(* Arrival Time Monitor core, an abstract base by convention: thin ND-framework
   state-mover wrapper that holds only references, interfaces and the shared
   sub-FBs. The state bridge is here as REFERENCE TO UINT (eEnumSetRef and
   eEnumGetRef) and the body runs on it, but the enum variables, the state
   storage and the state names belong to the derived type, which passes them
   in. Y mover via FB_PositionStatePMPSND over one motor, plus a
   tick site for the in-beam thermocouple and flow meter.

   A derived type supplies everything that depends on the state list:
     - eEnumSet and eEnumGet, the device enum (UINT base, OUT = 1, then the
       targets) with the MMS:STATE:SET and MMS:STATE:GET pytmc pragmas, so the
       EPICS state menu comes from that enum;
     - afbStateDefaults, one FB_CC_InternalStateConfig per state, which writes
       the per-state sName and fDelta;
     - an FB_Init that repeats the inputs below and binds eEnumSetRef and
       eEnumGetRef to the enum variables, and a CallAfterInit that calls the
       configurators. The base CallAfterInit runs on its own through the
       call_after_init attribute.
   FB_ATM is the library derived type (E_ATM_States). A device with another
   state list derives this FB the same way.

   State 1 is OUT, which vetoes the thermocouple. *)
{attribute 'call_after_init'}
FUNCTION_BLOCK FB_ATM_Core
VAR
    {attribute 'pytmc' := 'pv: STC:01'}
    fbTempSensor1 : FB_CC_TempSensor;

    {attribute 'pytmc' := 'pv: FWM'}
    fbFlowMeter : FB_AnalogInput := (iTermBits := 15, fTermMax := 60, fTermMin := 0);

    {attribute 'no_copy'}
    aiMotionStage         : REFERENCE TO ARRAY[1..MotionConstants.MAX_STATE_MOTORS] OF I_MotionStage;
    {attribute 'no_copy'}
    astPositionState      : REFERENCE TO ARRAY[1..MotionConstants.MAX_STATE_MOTORS]
                                            OF ARRAY[1..GeneralConstants.MAX_STATES] OF ST_PositionState;
    {attribute 'no_copy'}
    fbFFHWO               : REFERENCE TO FB_HardwareFFOutput;
    {attribute 'no_copy'}
    fbArbiter             : REFERENCE TO FB_Arbiter;
    sDeviceName           : STRING;
    sTransitionKey        : STRING;
    bEnableMotion         : BOOL := TRUE;
    bEnableBeamParams     : BOOL;
    bEnablePositionLimits : BOOL;
    bReadDBNow            : BOOL;
    bFileReaderBusy       : REFERENCE TO BOOL;
    bFileReaderError      : REFERENCE TO BOOL;

    {attribute 'no_copy'}
    eEnumSetRef           : REFERENCE TO UINT;
    {attribute 'no_copy'}
    eEnumGetRef           : REFERENCE TO UINT;

    {attribute 'pytmc' := 'pv: MMS'}
    fbStates : FB_PositionStatePMPSND(
        aiMotionStage         := aiMotionStage,
        astPositionState      := astPositionState,
        nActiveMotorCount     := nStateMotorCount,
        eEnumSet              := eEnumSetRef,
        eEnumGet              := eEnumGetRef,
        bEnableMotion         := bEnableMotion,
        eMotionRequestPolicy  := E_MotionRequestPolicy.INTERRUPT,
        bEnableBeamParams     := bEnableBeamParams,
        bEnablePositionLimits := bEnablePositionLimits,
        bReadDBNow            := bReadDBNow,
        bFileReaderBusy       := bFileReaderBusy,
        bFileReaderError      := bFileReaderError,
        fbFFHWO               := fbFFHWO,
        fbArbiter             := fbArbiter,
        sDeviceName           := sDeviceName,
        sTransitionKey        := sTransitionKey
    );
END_VAR
VAR_OUTPUT
    // The PMPS database lookup associated with the current position state.
    stDbStateParams: ST_DbStateParams;
END_VAR
VAR CONSTANT
    (* Number of motors the state mover drives. Every device here has one state
       motor, in slot 1; the code around fbStates assumes it. *)
    nStateMotorCount : UINT := 1;
    (* ATM-wide default tolerance for state in-position detection. Derived
       types pass it to their afbStateDefaults. *)
    FDELTA_DEFAULT : LREAL := 2;
    // State value of OUT in every ATM enum.
    nOutState : UINT := 1;
END_VAR

IF NOT __ISVALIDREF(aiMotionStage)
   OR NOT __ISVALIDREF(astPositionState)
   OR NOT __ISVALIDREF(fbFFHWO)
   OR NOT __ISVALIDREF(fbArbiter)
   OR NOT __ISVALIDREF(eEnumSetRef)
   OR NOT __ISVALIDREF(eEnumGetRef) THEN
    RETURN;
END_IF

fbStates(
    stDbStateParams => stDbStateParams
);

// Faults only while something is in the beam (not OUT).
fbTempSensor1(
    fFaultThreshold := fbStates.stDbStateParams.stReactiveParams.nTempSP,
    bVeto           := eEnumGetRef = nOutState,
    sDevName        := sDeviceName,
    io_fbFFHWO      := fbFFHWO
);

fbFlowMeter();

(* Auto-fired after FB_Init. Wires fbStates through CallAfterInitCore. *)
{attribute 'call_after_init'}
METHOD CallAfterInit
THIS^.CallAfterInitCore();
END_METHOD

(* Wires fbStates with the references this FB holds, through
   CallAfterInitStateMover / CallAfterInitPMPS, because fbStates' inline-init
   ran first and forwarded nil refs. Does nothing while the essential refs are
   still nil. CallAfterInit calls it. A derived type that was re-wired after its
   host FB's CallAfterInit calls it again through SUPER^. *)
METHOD CallAfterInitCore
IF NOT __ISVALIDREF(aiMotionStage)
   OR NOT __ISVALIDREF(astPositionState)
   OR NOT __ISVALIDREF(eEnumSetRef)
   OR NOT __ISVALIDREF(eEnumGetRef) THEN
    RETURN;
END_IF

THIS^.fbStates.CallAfterInitStateMover(
    aiMotionStage         := aiMotionStage,
    astPositionState      := astPositionState,
    nActiveMotorCount     := nStateMotorCount,
    eEnumSet              := eEnumSetRef,
    eEnumGet              := eEnumGetRef,
    bEnableMotion         := bEnableMotion,
    eMotionRequestPolicy  := E_MotionRequestPolicy.INTERRUPT,
);

THIS^.fbStates.CallAfterInitPMPS(
    aiMotionStage         := aiMotionStage,
    astPositionState      := astPositionState,
    bEnableBeamParams     := bEnableBeamParams,
    bEnablePositionLimits := bEnablePositionLimits,
    bReadDBNow            := bReadDBNow,
    bFileReaderBusy       := bFileReaderBusy,
    bFileReaderError      := bFileReaderError,
    fbFFHWO               := fbFFHWO,
    fbArbiter             := fbArbiter,
    sDeviceName           := sDeviceName,
    sTransitionKey        := sTransitionKey
);
END_METHOD

(* Stores FB_Init inputs into instance fields; every non-value input is
   REFERENCE TO, REF= bound for the FB lifetime. fbStates inline-init
   captured these params at construction, so this records the same refs
   on THIS^ for body use and live caller writes. *)
{attribute 'analysis' := '-33'}
METHOD FB_Init : BOOL
VAR_INPUT
    bInitRetains           : BOOL;
    bInCopyCode            : BOOL;
    aiMotionStage          : REFERENCE TO ARRAY[1..MotionConstants.MAX_STATE_MOTORS] OF I_MotionStage;
    astPositionState       : REFERENCE TO ARRAY[1..MotionConstants.MAX_STATE_MOTORS]
                                            OF ARRAY[1..GeneralConstants.MAX_STATES] OF ST_PositionState;
    fbFFHWO                : REFERENCE TO FB_HardwareFFOutput;
    fbArbiter              : REFERENCE TO FB_Arbiter;
    sDeviceName            : STRING;
    sTransitionKey         : STRING;
    bEnableBeamParams      : BOOL;
    bEnablePositionLimits  : BOOL;
    bReadDBNow             : BOOL;
    bFileReaderBusy        : REFERENCE TO BOOL;
    bFileReaderError       : REFERENCE TO BOOL;
END_VAR
THIS^.aiMotionStage    REF= aiMotionStage;
THIS^.astPositionState REF= astPositionState;
THIS^.fbFFHWO          REF= fbFFHWO;
THIS^.fbArbiter        REF= fbArbiter;
THIS^.sDeviceName      := sDeviceName;
THIS^.sTransitionKey   := sTransitionKey;
THIS^.bEnableBeamParams     := bEnableBeamParams;
THIS^.bEnablePositionLimits := bEnablePositionLimits;
THIS^.bReadDBNow            := bReadDBNow;
THIS^.bFileReaderBusy       REF= bFileReaderBusy;
THIS^.bFileReaderError      REF= bFileReaderError;
END_METHOD

END_FUNCTION_BLOCK

(* stored: Version 1.1.0.1
   POU FB_ATM_Core: Id {0b07f9bb-47d7-44ec-ac70-db2931ab90d6}, SpecialFunc None
   Method CallAfterInit: Id {a97fcae5-1420-4268-8023-befe115b659f}
   Method CallAfterInitCore: Id {85d661a7-6fb2-44c7-9a53-7e1119321676}
   Method FB_Init: Id {7eff5e72-784e-45c9-8b75-c8d832df35eb} *)
